// TIA Portal V20 export
// export: Created 2026-10-20T18:55:14.1957278Z, ExportSetting None, DisplayName Totally Integrated Automation Portal, DisplayVersion V20 Update 6, DisplayName TIA Portal Openness, DisplayVersion V20 Update 6, DisplayName TIA Portal Version Control Interface, DisplayVersion V20 Update 6, DisplayName SINAMICS Startdrive Advanced, DisplayVersion V20 SP1, DisplayName SINAMICS Startdrive G130, G150, S120, S150, SINAMICS MV, G220, S200, S210, DisplayVersion V20 SP1, DisplayName SINAMICS Startdrive G110M, G120, G120C, G120D, G120P, G115D, DisplayVersion V20 SP1, DisplayName STEP 7 Professional, DisplayVersion V20 Update 6, DisplayName STEP 7 Safety, DisplayVersion V20 Update 2, DisplayName WinCC Basic/Comfort/Advanced, DisplayVersion V20 Update 6, DisplayName WinCC Unified, DisplayVersion V20 Update 6
VAR_GLOBAL   // PLC tag table "IO_Remote_Panel_4"
   "VTD4 PUSH TO ENTER VTD ZONE" AT %I1053.4 : Bool;
   "STO VTD - CH2(4)" AT %Q1081.1 : Bool;
   "CABINET COOLING FAN CIRCUIT BREAKER FEEDBACK(4)" AT %I1055.3 : Bool;
   "VTD4 UPPER LIMIT" AT %I1052.0 : Bool;
   "STO CNV VFD (Level 4,5,6 - Side1) - CH2(4)" AT %Q1081.7 : Bool;
   "STO CNV VFD (Level 1,2,3 - Side1) - CH1(4)" AT %Q1081.4 : Bool;
   "C4102_SFTY STOPPER ROTATE" AT %Q505.4 : Bool;
   "Power Enable Safety Stopper Conveyors (Level 4,5,6 - Side1) - CH1(4)" AT %Q1093.2 : Bool;
   "C4108_SFTY STOPPER ROTATE" AT %Q513.4 : Bool;
   "Chain Slack 3 - CH1(4)" AT %I1067.2 : Bool;   // Chain Slack 3 - CH1
   "Chain Slack 2 - CH1(4)" AT %I1067.1 : Bool;   // Chain Slack 2 - CH1
   "SCA 4001 STACK LIGHTS YELLOW" AT %Q519.5 : Bool;
   "STO CNV VFD (Level 7,8 - Side1) - CH2(4)" AT %Q1087.1 : Bool;
   "VTU HOIST BRAKE SAFETY ENABLE 1(4)" AT %Q1093.6 : Bool;
   "C4107_SFTY STOPPER ROTATE" AT %Q513.0 : Bool;
   "VTU HOIST BRAKE SAFETY ENABLE EDM FEEDBACK(4)" AT %I1074.3 : Bool;
   "Chain Slack 3 - CH2(4)" AT %I1067.6 : Bool;   // Chain Slack 3 - CH2
   "C4107 CIRCUIT BREAKER FEEDBACK" AT %I1054.6 : Bool;
   "VTD4 SFTY STOPPER CNVS 7,8 - (SIDE 1)" AT %I1074.2 : Bool;
   "CABINET 24V PSU CIRCUIT BREAKER FEEDBACK(4)" AT %I1055.2 : Bool;
   "Power Enable Safety Stopper Conveyors (Level 7,8 - Side1) - CH2(4)" AT %Q1093.5 : Bool;
   "Power Enable Safety Stopper Conveyors (Level 1,2,3 - Side1) - CH1(4)" AT %Q1093.0 : Bool;
   "C4106 CIRCUIT BREAKER FEEDBACK" AT %I1054.5 : Bool;
   "STO VTD - CH1(4)" AT %Q1081.0 : Bool;
   "C4103 CIRCUIT BREAKER FEEDBACK" AT %I1054.2 : Bool;
   "VTD4 CIRCUIT BREAKER FEEDBACK" AT %I1055.1 : Bool;
   "VTU HOIST BRAKE SAFETY ENABLE 2(4)" AT %Q1093.7 : Bool;
   "C4103_SFTY STOPPER ROTATE" AT %Q506.0 : Bool;
   "Power Enable Safety Stopper Conveyors (Level 1,2,3 - Side1) - CH2(4)" AT %Q1093.1 : Bool;
   "RESET (CABINET)(4)" AT %I1060.3 : Bool;   // Reset (Cabinet) - CH1
   "STO CNV VFD (Level 4,5,6 - Side1) - CH1(4)" AT %Q1081.6 : Bool;
   "VTD4 PUSH TO EXIT VTD ZONE" AT %I1053.5 : Bool;
   "C4104_SFTY STOPPER ROTATE" AT %Q506.4 : Bool;
   "Power Enable Safety Stopper Conveyors (Level 4,5,6 - Side1) - CH2(4)" AT %Q1093.3 : Bool;
   "C4101_SFTY STOPPER ROTATE" AT %Q505.0 : Bool;
   "STO CNV VFD (Level 1,2,3 - Side1) - CH2(4)" AT %Q1081.5 : Bool;
   "STO CONVEYOR VTD - CH1(4)" AT %Q1081.2 : Bool;
   "OVERTRAVEL UPPER LIMIT - CH1(4)" AT %I1060.1 : Bool;   // Overtravel Upper Limit - CH1
   "STO CONVEYOR VTD - CH2(4)" AT %Q1081.3 : Bool;
   "C4105 CIRCUIT BREAKER FEEDBACK" AT %I1054.4 : Bool;
   "Chain Slack 4 - CH1(4)" AT %I1067.3 : Bool;   // Chain Slack 4 - CH1
   "Chain Slack 1 - CH1(4)" AT %I1067.0 : Bool;   // Chain Slack 1 - CH1
   "C4102 CIRCUIT BREAKER FEEDBACK" AT %I1054.1 : Bool;
   "C4108 CIRCUIT BREAKER FEEDBACK" AT %I1054.7 : Bool;
   "VTD4 LOWER LIMIT" AT %I1052.3 : Bool;
   "OVERTRAVEL LOWER LIMIT - CH1(4)" AT %I1060.0 : Bool;   // Overtravel Lower Limit - CH1
   "E-STOP (CABINET) - CH1(4)" AT %I1060.2 : Bool;   // E-Stop (Cabinet)- CH1
   "CVTD4 CIRCUIT BREAKER FEEDBACK" AT %I1055.0 : Bool;
   "C4101 CIRCUIT BREAKER FEEDBACK" AT %I1054.0 : Bool;
   "OVERTRAVEL LOWER LIMIT - CH2(4)" AT %I1060.4 : Bool;   // Overtravel Lower Limit - CH2
   "VTD4 SFTY STOPPER CNVS 1,2,3 - (SIDE 1)" AT %I1074.0 : Bool;   // SAFETY STOPPER CONVEYORS (1,2,3 - SIDE 1) EDMFEEDBACK
   "C4104 CIRCUIT BREAKER FEEDBACK" AT %I1054.3 : Bool;
   "C4106_SFTY STOPPER ROTATE" AT %Q512.4 : Bool;
   "EMERGENCY STOP RESET STATUS - ON(4)" AT %Q520.4 : Bool;   // 920SL1
   "C4105_SFTY STOPPER ROTATE" AT %Q512.0 : Bool;
   "Chain Slack 1 - CH2(4)" AT %I1067.4 : Bool;   // Chain Slack 1 - CH2
   "STO CNV VFD (Level 7,8 - Side1) - CH1(4)" AT %Q1087.0 : Bool;
   "OVERTRAVEL UPPER LIMIT - CH2(4)" AT %I1060.5 : Bool;   // Overtravel Upper Limit - CH2
   "Power Enable Safety Stopper Conveyors (Level 7,8 - Side1) - CH1(4)" AT %Q1093.4 : Bool;
   "Chain Slack 4 - CH2(4)" AT %I1067.7 : Bool;   // Chain Slack 4 - CH2
   "Chain Slack 2 - CH2(4)" AT %I1067.5 : Bool;   // Chain Slack 2 - CH2
   "E-STOP (CABINET) - CH2(4)" AT %I1060.6 : Bool;   // E-Stop (Cabinet) - CH2
   "SCA 4001 STACK LIGHTS GREEN" AT %Q519.6 : Bool;
   "SCA 4001 STACK LIGHTS RED" AT %Q519.4 : Bool;
   "VTD4 DOCKING PINS 1 EXTEND" AT %Q520.2 : Bool;
   "VTD4 DOCKING PINS 2 EXTEND" AT %Q520.0 : Bool;
   "VTD4 DOCKING PINS 2 RETRACT" AT %Q520.1 : Bool;
   "VTD4 DOCKING PINS 1 RETRACT" AT %Q520.3 : Bool;
   "GATE_SENSOR_CH2(4)" AT %I1074.5 : Bool;
   "VTD4 SFTY STOPPER CNVS 4,5,6 - (SIDE 1)" AT %I1074.4 : Bool;
   "GATE_SENSOR_CH1(4)" AT %I1074.1 : Bool;
END_VAR
